// TIA Portal V19 export
TYPE "EM06_Input"
   STRUCT
      Cmds { S7_SetPoint := 'True'} : "EM_Input";
      CtrlMode : Int;   // 0=Off, 1=Descarga de masa, 2=Desague de lavado
      NivelDescargaOn : Real;   // Nivel del recibidor para iniciar descarga
      NivelDescargaOff : Real;   // Nivel del recibidor para pausar descarga
      NivelDescargaFin : Real;   // Nivel de tacho considerado vacio
      EmptyFilter : Time;   // Permanencia bajo nivel de fin para completar
      DrainTime : Time;   // Tiempo de apertura del desague
      VacuumBrokenPermit : Bool;   // Permiso para descargar masa con vacio roto
   END_STRUCT;
END_TYPE
